FUNCTION_BLOCK TestFb
VAR_INPUT
	    stIn            : ST_NordSK550P_In;
END_VAR
VAR_OUTPUT
	    wStatusWord      : UINT;
		dupa2 : INT;
END_VAR
VAR
	dupa : INT := 100;
	i : INT;
END_VAR

wStatusWord := stIn.wStatusWord;
dupa := dupa2;

END_FUNCTION_BLOCK

(* stored: Version 1.1.0.1
   POU TestFb: Id {7ffda057-922e-4c73-8527-4d253acdd599}, SpecialFunc None *)
